Staubli VAL3: unLock.pgx

program unLock()
  local string l_sEntry
  local bool l_bResult
  local num i
begin
//  if bLock==true
//    l_bResult=userPagePrompt("请输入密码",l_sEntry)
//    if l_bResult==false
//      return
//    endIf
//    if l_sEntry!=sPassword[0]
//      popUpMsg("密码错误")
//      return
//    endIf
//    //2024.04.29 add解锁扭矩限位设置
//    for i=0 to size(bDisable)-1
//      bDisable[i]=false
//    endFor
//    popUpMsg("修改后请点击保存!")
//    bLock=false
//  else
//    for i=0 to size(bDisable)-1
//      bDisable[i]=true
//    endFor
//    call seMaxJntForce()
//    call libTqe:_getSetForce(nMaxJntForec)
//    popUpMsg("机器人关节扭矩限制保存成功!")
//    bLock=true
//  endIf
end
